(* IEC 61131-3 sources: codesys-framework/txt/application/WeVe Core (library)/00 Application/FB_Application, 1 file *)

(* ---- InitializeEvents.method.st ---- *)
METHOD PROTECTED ABSTRACT InitializeEvents : BOOL
VAR_INPUT
END_VAR
